(*

**Numerical footnote**

Footnote references, like [5]_. Note that footnotes may get rearranged, e.g., to the bottom of the "page".

--------

.. [5] A numerical footnote. Note there's no colon after the ``]``.
*)

FUNCTION_BLOCK FB_Libdoc_ManuallyNumberedFootnotes
VAR_INPUT
    nVarA : INT;
    nVarB : INT;
END_VAR
VAR_OUTPUT
    nSum : INT;
END_VAR
VAR
END_VAR

END_FUNCTION_BLOCK

(* stored: Version 1.1.0.1, ProductVersion 3.1.4022.17
   POU FB_Libdoc_ManuallyNumberedFootnotes: Id {2611b9ed-1882-4766-bc40-e4e3dead1038}, SpecialFunc None *)
